(* IEC 61131-3 sources: 2026_Projet_YGO_ExcavatriceDragage/TOOLS/TEST_AUTO_CI/RESULTS/B_AU_SECURITE/tests/contract_deferred, 1 file *)

(* ---- test_fb_safety_emergency_contract_deferred.st ---- *)
(* Essais différés : causes, diagnostics et latches. Non exécutés par run.bat ; à reprendre dans le futur socle de contrat FB. *)
SETUP
VAR
    fb : FB_SAFETY_EMERGENCYMANAGEMENT;
END_VAR
END_SETUP

(* Ce fichier est volontairement hors execution run.bat. Migration prevue vers le socle de contrat FB. *)

TEST 'TC-P01-023 Etape invalide -> abandon trace et lockout'
    fb(ENABLE := TRUE, RESET := FALSE, ARMREQUEST := FALSE, POWERCUTOFFREQUEST := FALSE,
       BTNEMERGENCYCUTOFF := FALSE, EMERGENCYCHAINCLOSED := TRUE, POWERCONTACTORENGAGED := FALSE);
    fb(ENABLE := TRUE, RESET := FALSE, ARMREQUEST := FALSE, POWERCUTOFFREQUEST := FALSE,
       BTNEMERGENCYCUTOFF := FALSE, EMERGENCYCHAINCLOSED := TRUE, POWERCONTACTORENGAGED := FALSE);

    fb.ARMINGSEQSTEP := 7;
    ADVANCE_TIME(10000000);
    fb(ENABLE := TRUE, RESET := FALSE, ARMREQUEST := FALSE, POWERCUTOFFREQUEST := FALSE,
       BTNEMERGENCYCUTOFF := FALSE, EMERGENCYCHAINCLOSED := TRUE, POWERCONTACTORENGAGED := FALSE);
    fb(ENABLE := TRUE, RESET := FALSE, ARMREQUEST := FALSE, POWERCUTOFFREQUEST := FALSE,
       BTNEMERGENCYCUTOFF := FALSE, EMERGENCYCHAINCLOSED := TRUE, POWERCONTACTORENGAGED := FALSE);

    ASSERT_EQ(fb.STATUS.STATE.STEP, 0, 'etape inconnue -> IDLE');
    ASSERT_EQ(fb.STATUS.DIAG.LASTABORTSTEP, 7, 'etape inconnue tracee');
    ASSERT_EQ(fb.STATUS.DIAG.LASTABORTCAUSE, 256, 'cause = CST_ABORT_INVALID_STEP');
    ASSERT_TRUE(fb.STATUS.DIAG.LOCKOUTACTIVE, 'etape inconnue -> lockout');
    ASSERT_FALSE(fb.CMD.ARMPULSE_CMD, 'etape inconnue -> aucune impulsion');
    ASSERT_EQ(fb.STATUS.OPERATORMESSAGE, 'AU: etape sequence invalide - verifier puis Reset', 'etape inconnue -> message explicite');
END_TEST

TEST 'TC-P01-011 PowerCutOffRequest pendant l impulsion (step 5) -> abandon 16#0010 + lockout + Error=FALSE'
    (* Montee nominale jusqu au pulse (step 5), comme TC-P01-003 *)
    fb(ENABLE := TRUE, RESET := FALSE, ARMREQUEST := FALSE, POWERCUTOFFREQUEST := FALSE,
       BTNEMERGENCYCUTOFF := FALSE, EMERGENCYCHAINCLOSED := TRUE, POWERCONTACTORENGAGED := FALSE);
    fb(ENABLE := TRUE, RESET := FALSE, ARMREQUEST := FALSE, POWERCUTOFFREQUEST := FALSE,
       BTNEMERGENCYCUTOFF := FALSE, EMERGENCYCHAINCLOSED := TRUE, POWERCONTACTORENGAGED := FALSE);
    ADVANCE_TIME(10000000);
    fb(ENABLE := TRUE, RESET := FALSE, ARMREQUEST := FALSE, POWERCUTOFFREQUEST := FALSE,
       BTNEMERGENCYCUTOFF := FALSE, EMERGENCYCHAINCLOSED := TRUE, POWERCONTACTORENGAGED := FALSE);
    fb(ENABLE := TRUE, RESET := FALSE, ARMREQUEST := FALSE, POWERCUTOFFREQUEST := FALSE,
       BTNEMERGENCYCUTOFF := FALSE, EMERGENCYCHAINCLOSED := TRUE, POWERCONTACTORENGAGED := FALSE);
    ADVANCE_TIME(10000000);
    fb(ENABLE := TRUE, RESET := FALSE, ARMREQUEST := TRUE, POWERCUTOFFREQUEST := FALSE,
       BTNEMERGENCYCUTOFF := FALSE, EMERGENCYCHAINCLOSED := TRUE, POWERCONTACTORENGAGED := FALSE);
    fb(ENABLE := TRUE, RESET := FALSE, ARMREQUEST := TRUE, POWERCUTOFFREQUEST := FALSE,
       BTNEMERGENCYCUTOFF := FALSE, EMERGENCYCHAINCLOSED := TRUE, POWERCONTACTORENGAGED := FALSE);
    ADVANCE_TIME(200000000);
    fb(ENABLE := TRUE, RESET := FALSE, ARMREQUEST := FALSE, POWERCUTOFFREQUEST := FALSE,
       BTNEMERGENCYCUTOFF := FALSE, EMERGENCYCHAINCLOSED := FALSE, POWERCONTACTORENGAGED := FALSE);
    fb(ENABLE := TRUE, RESET := FALSE, ARMREQUEST := FALSE, POWERCUTOFFREQUEST := FALSE,
       BTNEMERGENCYCUTOFF := FALSE, EMERGENCYCHAINCLOSED := FALSE, POWERCONTACTORENGAGED := FALSE);
    ADVANCE_TIME(200000000);
    fb(ENABLE := TRUE, RESET := FALSE, ARMREQUEST := FALSE, POWERCUTOFFREQUEST := FALSE,
       BTNEMERGENCYCUTOFF := FALSE, EMERGENCYCHAINCLOSED := TRUE, POWERCONTACTORENGAGED := FALSE);
    fb(ENABLE := TRUE, RESET := FALSE, ARMREQUEST := FALSE, POWERCUTOFFREQUEST := FALSE,
       BTNEMERGENCYCUTOFF := FALSE, EMERGENCYCHAINCLOSED := TRUE, POWERCONTACTORENGAGED := FALSE);
    ADVANCE_TIME(200000000);
    fb(ENABLE := TRUE, RESET := FALSE, ARMREQUEST := FALSE, POWERCUTOFFREQUEST := FALSE,
       BTNEMERGENCYCUTOFF := FALSE, EMERGENCYCHAINCLOSED := FALSE, POWERCONTACTORENGAGED := FALSE);
    fb(ENABLE := TRUE, RESET := FALSE, ARMREQUEST := FALSE, POWERCUTOFFREQUEST := FALSE,
       BTNEMERGENCYCUTOFF := FALSE, EMERGENCYCHAINCLOSED := FALSE, POWERCONTACTORENGAGED := FALSE);
    ADVANCE_TIME(200000000);
    fb(ENABLE := TRUE, RESET := FALSE, ARMREQUEST := FALSE, POWERCUTOFFREQUEST := FALSE,
       BTNEMERGENCYCUTOFF := FALSE, EMERGENCYCHAINCLOSED := TRUE, POWERCONTACTORENGAGED := FALSE);
    fb(ENABLE := TRUE, RESET := FALSE, ARMREQUEST := FALSE, POWERCUTOFFREQUEST := FALSE,
       BTNEMERGENCYCUTOFF := FALSE, EMERGENCYCHAINCLOSED := TRUE, POWERCONTACTORENGAGED := FALSE);
    ASSERT_EQ(fb.STATUS.STATE.STEP, 5, 'les 2 canaux valides -> pulse (step 5)');
    ASSERT_TRUE(fb.CMD.ARMPULSE_CMD, 'precondition : pulse actif');

    (* Coupure metier PowerCutOffRequest PENDANT l impulsion (step 5) *)
    ADVANCE_TIME(10000000);
    fb(ENABLE := TRUE, RESET := FALSE, ARMREQUEST := FALSE, POWERCUTOFFREQUEST := TRUE,
       BTNEMERGENCYCUTOFF := FALSE, EMERGENCYCHAINCLOSED := TRUE, POWERCONTACTORENGAGED := FALSE);
    fb(ENABLE := TRUE, RESET := FALSE, ARMREQUEST := FALSE, POWERCUTOFFREQUEST := TRUE,
       BTNEMERGENCYCUTOFF := FALSE, EMERGENCYCHAINCLOSED := TRUE, POWERCONTACTORENGAGED := FALSE);
    ASSERT_EQ(fb.STATUS.STATE.STEP, 0, 'PowerCutOff pendant pulse -> sequence ramenee a IDLE');
    ASSERT_EQ(fb.STATUS.DIAG.LASTABORTCAUSE, 16#0010, 'cause abandon = 16#0010 (PowerCutOff metier)');
    ASSERT_EQ(fb.STATUS.DIAG.LASTABORTSTEP, 5, 'abandon a l etape 5 (impulsion)');
    ASSERT_TRUE(fb.STATUS.DIAG.LOCKOUTACTIVE, 'lockout 5s actif apres coupure metier');
    ASSERT_FALSE(fb.STATUS.DIAG.ERROR, 'coupure metier voulue -> PAS de defaut d armement (Error=FALSE)');
    ASSERT_FALSE(fb.STATUS.STATE.ARMABLE, 'interlock : PowerCutOffRequest actif -> Armable=FALSE');
    ASSERT_EQ(fb.STATUS.OPERATORMESSAGE, 'AU: coupure securite metier active - lever la cause puis rearmer', 'message coupure metier (priorite §11 sur le CASE)');
END_TEST

TEST 'TC-P01-012 Armable=1 mais rearmement echoue a l etape 5 (PowerCutOff pendant pulse)'
    (* Precondition : au repos boucle saine, Armable=TRUE (rearmement autorise) *)
    fb(ENABLE := TRUE, RESET := FALSE, ARMREQUEST := FALSE, POWERCUTOFFREQUEST := FALSE,
       BTNEMERGENCYCUTOFF := FALSE, EMERGENCYCHAINCLOSED := TRUE, POWERCONTACTORENGAGED := FALSE);
    fb(ENABLE := TRUE, RESET := FALSE, ARMREQUEST := FALSE, POWERCUTOFFREQUEST := FALSE,
       BTNEMERGENCYCUTOFF := FALSE, EMERGENCYCHAINCLOSED := TRUE, POWERCONTACTORENGAGED := FALSE);
    ADVANCE_TIME(10000000);
    fb(ENABLE := TRUE, RESET := FALSE, ARMREQUEST := FALSE, POWERCUTOFFREQUEST := FALSE,
       BTNEMERGENCYCUTOFF := FALSE, EMERGENCYCHAINCLOSED := TRUE, POWERCONTACTORENGAGED := FALSE);
    fb(ENABLE := TRUE, RESET := FALSE, ARMREQUEST := FALSE, POWERCUTOFFREQUEST := FALSE,
       BTNEMERGENCYCUTOFF := FALSE, EMERGENCYCHAINCLOSED := TRUE, POWERCONTACTORENGAGED := FALSE);
    ASSERT_TRUE(fb.STATUS.STATE.ARMABLE, 'precondition : Armable=TRUE (rearmement autorise)');

    (* Rearmement lance -> sequence demarre *)
    ADVANCE_TIME(10000000);
    fb(ENABLE := TRUE, RESET := FALSE, ARMREQUEST := TRUE, POWERCUTOFFREQUEST := FALSE,
       BTNEMERGENCYCUTOFF := FALSE, EMERGENCYCHAINCLOSED := TRUE, POWERCONTACTORENGAGED := FALSE);
    fb(ENABLE := TRUE, RESET := FALSE, ARMREQUEST := TRUE, POWERCUTOFFREQUEST := FALSE,
       BTNEMERGENCYCUTOFF := FALSE, EMERGENCYCHAINCLOSED := TRUE, POWERCONTACTORENGAGED := FALSE);
    ASSERT_EQ(fb.STATUS.STATE.STEP, 1, 'ArmRequest -> sequence lancee (step 1)');

    (* Montee nominale jusqu au pulse (step 5) *)
    ADVANCE_TIME(200000000);
    fb(ENABLE := TRUE, RESET := FALSE, ARMREQUEST := FALSE, POWERCUTOFFREQUEST := FALSE,
       BTNEMERGENCYCUTOFF := FALSE, EMERGENCYCHAINCLOSED := FALSE, POWERCONTACTORENGAGED := FALSE);
    fb(ENABLE := TRUE, RESET := FALSE, ARMREQUEST := FALSE, POWERCUTOFFREQUEST := FALSE,
       BTNEMERGENCYCUTOFF := FALSE, EMERGENCYCHAINCLOSED := FALSE, POWERCONTACTORENGAGED := FALSE);
    ADVANCE_TIME(200000000);
    fb(ENABLE := TRUE, RESET := FALSE, ARMREQUEST := FALSE, POWERCUTOFFREQUEST := FALSE,
       BTNEMERGENCYCUTOFF := FALSE, EMERGENCYCHAINCLOSED := TRUE, POWERCONTACTORENGAGED := FALSE);
    fb(ENABLE := TRUE, RESET := FALSE, ARMREQUEST := FALSE, POWERCUTOFFREQUEST := FALSE,
       BTNEMERGENCYCUTOFF := FALSE, EMERGENCYCHAINCLOSED := TRUE, POWERCONTACTORENGAGED := FALSE);
    ADVANCE_TIME(200000000);
    fb(ENABLE := TRUE, RESET := FALSE, ARMREQUEST := FALSE, POWERCUTOFFREQUEST := FALSE,
       BTNEMERGENCYCUTOFF := FALSE, EMERGENCYCHAINCLOSED := FALSE, POWERCONTACTORENGAGED := FALSE);
    fb(ENABLE := TRUE, RESET := FALSE, ARMREQUEST := FALSE, POWERCUTOFFREQUEST := FALSE,
       BTNEMERGENCYCUTOFF := FALSE, EMERGENCYCHAINCLOSED := FALSE, POWERCONTACTORENGAGED := FALSE);
    ADVANCE_TIME(200000000);
    fb(ENABLE := TRUE, RESET := FALSE, ARMREQUEST := FALSE, POWERCUTOFFREQUEST := FALSE,
       BTNEMERGENCYCUTOFF := FALSE, EMERGENCYCHAINCLOSED := TRUE, POWERCONTACTORENGAGED := FALSE);
    fb(ENABLE := TRUE, RESET := FALSE, ARMREQUEST := FALSE, POWERCUTOFFREQUEST := FALSE,
       BTNEMERGENCYCUTOFF := FALSE, EMERGENCYCHAINCLOSED := TRUE, POWERCONTACTORENGAGED := FALSE);
    ASSERT_EQ(fb.STATUS.STATE.STEP, 5, 'les 2 canaux valides -> pulse (step 5)');

    (* Coupure metier pendant l impulsion -> echec a l etape 5 *)
    ADVANCE_TIME(10000000);
    fb(ENABLE := TRUE, RESET := FALSE, ARMREQUEST := FALSE, POWERCUTOFFREQUEST := TRUE,
       BTNEMERGENCYCUTOFF := FALSE, EMERGENCYCHAINCLOSED := TRUE, POWERCONTACTORENGAGED := FALSE);
    fb(ENABLE := TRUE, RESET := FALSE, ARMREQUEST := FALSE, POWERCUTOFFREQUEST := TRUE,
       BTNEMERGENCYCUTOFF := FALSE, EMERGENCYCHAINCLOSED := TRUE, POWERCONTACTORENGAGED := FALSE);
    ASSERT_EQ(fb.STATUS.STATE.STEP, 0, 'echec a l etape 5 -> sequence ramenee a IDLE');
    ASSERT_EQ(fb.STATUS.DIAG.LASTABORTSTEP, 5, 'abandon a l etape 5');
    ASSERT_EQ(fb.STATUS.DIAG.LASTABORTCAUSE, 16#0010, 'cause = 16#0010 (PowerCutOff metier)');
    ASSERT_FALSE(fb.STATUS.DONE, 'rearmement NON abouti (Done=FALSE, contacteur non engage)');
    ASSERT_FALSE(fb.STATUS.DIAG.ERROR, 'echec silencieux : PAS de defaut d armement (Error=FALSE)');
END_TEST

TEST 'TC-P01-013 Recuperation Reset : cause latched -> Reset -> cause levee -> rearmement reussi'
    (* Montee nominale jusqu au pulse (step 5), puis coupure metier -> abandon 16#0010 + lockout *)
    fb(ENABLE := TRUE, RESET := FALSE, ARMREQUEST := FALSE, POWERCUTOFFREQUEST := FALSE,
       BTNEMERGENCYCUTOFF := FALSE, EMERGENCYCHAINCLOSED := TRUE, POWERCONTACTORENGAGED := FALSE);
    fb(ENABLE := TRUE, RESET := FALSE, ARMREQUEST := FALSE, POWERCUTOFFREQUEST := FALSE,
       BTNEMERGENCYCUTOFF := FALSE, EMERGENCYCHAINCLOSED := TRUE, POWERCONTACTORENGAGED := FALSE);
    ADVANCE_TIME(10000000);
    fb(ENABLE := TRUE, RESET := FALSE, ARMREQUEST := FALSE, POWERCUTOFFREQUEST := FALSE,
       BTNEMERGENCYCUTOFF := FALSE, EMERGENCYCHAINCLOSED := TRUE, POWERCONTACTORENGAGED := FALSE);
    fb(ENABLE := TRUE, RESET := FALSE, ARMREQUEST := FALSE, POWERCUTOFFREQUEST := FALSE,
       BTNEMERGENCYCUTOFF := FALSE, EMERGENCYCHAINCLOSED := TRUE, POWERCONTACTORENGAGED := FALSE);
    ADVANCE_TIME(10000000);
    fb(ENABLE := TRUE, RESET := FALSE, ARMREQUEST := TRUE, POWERCUTOFFREQUEST := FALSE,
       BTNEMERGENCYCUTOFF := FALSE, EMERGENCYCHAINCLOSED := TRUE, POWERCONTACTORENGAGED := FALSE);
    fb(ENABLE := TRUE, RESET := FALSE, ARMREQUEST := TRUE, POWERCUTOFFREQUEST := FALSE,
       BTNEMERGENCYCUTOFF := FALSE, EMERGENCYCHAINCLOSED := TRUE, POWERCONTACTORENGAGED := FALSE);
    ADVANCE_TIME(200000000);
    fb(ENABLE := TRUE, RESET := FALSE, ARMREQUEST := FALSE, POWERCUTOFFREQUEST := FALSE,
       BTNEMERGENCYCUTOFF := FALSE, EMERGENCYCHAINCLOSED := FALSE, POWERCONTACTORENGAGED := FALSE);
    fb(ENABLE := TRUE, RESET := FALSE, ARMREQUEST := FALSE, POWERCUTOFFREQUEST := FALSE,
       BTNEMERGENCYCUTOFF := FALSE, EMERGENCYCHAINCLOSED := FALSE, POWERCONTACTORENGAGED := FALSE);
    ADVANCE_TIME(200000000);
    fb(ENABLE := TRUE, RESET := FALSE, ARMREQUEST := FALSE, POWERCUTOFFREQUEST := FALSE,
       BTNEMERGENCYCUTOFF := FALSE, EMERGENCYCHAINCLOSED := TRUE, POWERCONTACTORENGAGED := FALSE);
    fb(ENABLE := TRUE, RESET := FALSE, ARMREQUEST := FALSE, POWERCUTOFFREQUEST := FALSE,
       BTNEMERGENCYCUTOFF := FALSE, EMERGENCYCHAINCLOSED := TRUE, POWERCONTACTORENGAGED := FALSE);
    ADVANCE_TIME(200000000);
    fb(ENABLE := TRUE, RESET := FALSE, ARMREQUEST := FALSE, POWERCUTOFFREQUEST := FALSE,
       BTNEMERGENCYCUTOFF := FALSE, EMERGENCYCHAINCLOSED := FALSE, POWERCONTACTORENGAGED := FALSE);
    fb(ENABLE := TRUE, RESET := FALSE, ARMREQUEST := FALSE, POWERCUTOFFREQUEST := FALSE,
       BTNEMERGENCYCUTOFF := FALSE, EMERGENCYCHAINCLOSED := FALSE, POWERCONTACTORENGAGED := FALSE);
    ADVANCE_TIME(200000000);
    fb(ENABLE := TRUE, RESET := FALSE, ARMREQUEST := FALSE, POWERCUTOFFREQUEST := FALSE,
       BTNEMERGENCYCUTOFF := FALSE, EMERGENCYCHAINCLOSED := TRUE, POWERCONTACTORENGAGED := FALSE);
    fb(ENABLE := TRUE, RESET := FALSE, ARMREQUEST := FALSE, POWERCUTOFFREQUEST := FALSE,
       BTNEMERGENCYCUTOFF := FALSE, EMERGENCYCHAINCLOSED := TRUE, POWERCONTACTORENGAGED := FALSE);
    ASSERT_EQ(fb.STATUS.STATE.STEP, 5, 'pulse (step 5)');

    (* Coupure metier -> abandon 16#0010 + lockout *)
    ADVANCE_TIME(10000000);
    fb(ENABLE := TRUE, RESET := FALSE, ARMREQUEST := FALSE, POWERCUTOFFREQUEST := TRUE,
       BTNEMERGENCYCUTOFF := FALSE, EMERGENCYCHAINCLOSED := TRUE, POWERCONTACTORENGAGED := FALSE);
    fb(ENABLE := TRUE, RESET := FALSE, ARMREQUEST := FALSE, POWERCUTOFFREQUEST := TRUE,
       BTNEMERGENCYCUTOFF := FALSE, EMERGENCYCHAINCLOSED := TRUE, POWERCONTACTORENGAGED := FALSE);
    ASSERT_EQ(fb.STATUS.DIAG.LASTABORTCAUSE, 16#0010, 'cause latched = 16#0010');
    ASSERT_TRUE(fb.STATUS.DIAG.LOCKOUTACTIVE, 'lockout actif');

    (* Cause levee (PowerCutOffRequest=FALSE) + Reset -> lockout purge, Armable redevient TRUE *)
    ADVANCE_TIME(10000000);
    fb(ENABLE := TRUE, RESET := TRUE, ARMREQUEST := FALSE, POWERCUTOFFREQUEST := FALSE,
       BTNEMERGENCYCUTOFF := FALSE, EMERGENCYCHAINCLOSED := TRUE, POWERCONTACTORENGAGED := FALSE);
    fb(ENABLE := TRUE, RESET := TRUE, ARMREQUEST := FALSE, POWERCUTOFFREQUEST := FALSE,
       BTNEMERGENCYCUTOFF := FALSE, EMERGENCYCHAINCLOSED := TRUE, POWERCONTACTORENGAGED := FALSE);
    ASSERT_FALSE(fb.STATUS.DIAG.LOCKOUTACTIVE, 'Reset purge le lockout');
    ASSERT_TRUE(fb.STATUS.STATE.ARMABLE, 'cause levee + Reset -> Armable=TRUE');

    (* Nouveau rearmement -> reussite (contacteur engage) *)
    ADVANCE_TIME(10000000);
    fb(ENABLE := TRUE, RESET := FALSE, ARMREQUEST := TRUE, POWERCUTOFFREQUEST := FALSE,
       BTNEMERGENCYCUTOFF := FALSE, EMERGENCYCHAINCLOSED := TRUE, POWERCONTACTORENGAGED := FALSE);
    fb(ENABLE := TRUE, RESET := FALSE, ARMREQUEST := TRUE, POWERCUTOFFREQUEST := FALSE,
       BTNEMERGENCYCUTOFF := FALSE, EMERGENCYCHAINCLOSED := TRUE, POWERCONTACTORENGAGED := FALSE);
    ASSERT_EQ(fb.STATUS.STATE.STEP, 1, 'nouveau front ArmRequest -> sequence relancee');
    ADVANCE_TIME(200000000);
    fb(ENABLE := TRUE, RESET := FALSE, ARMREQUEST := FALSE, POWERCUTOFFREQUEST := FALSE,
       BTNEMERGENCYCUTOFF := FALSE, EMERGENCYCHAINCLOSED := FALSE, POWERCONTACTORENGAGED := FALSE);
    fb(ENABLE := TRUE, RESET := FALSE, ARMREQUEST := FALSE, POWERCUTOFFREQUEST := FALSE,
       BTNEMERGENCYCUTOFF := FALSE, EMERGENCYCHAINCLOSED := FALSE, POWERCONTACTORENGAGED := FALSE);
    ADVANCE_TIME(200000000);
    fb(ENABLE := TRUE, RESET := FALSE, ARMREQUEST := FALSE, POWERCUTOFFREQUEST := FALSE,
       BTNEMERGENCYCUTOFF := FALSE, EMERGENCYCHAINCLOSED := TRUE, POWERCONTACTORENGAGED := FALSE);
    fb(ENABLE := TRUE, RESET := FALSE, ARMREQUEST := FALSE, POWERCUTOFFREQUEST := FALSE,
       BTNEMERGENCYCUTOFF := FALSE, EMERGENCYCHAINCLOSED := TRUE, POWERCONTACTORENGAGED := FALSE);
    ADVANCE_TIME(200000000);
    fb(ENABLE := TRUE, RESET := FALSE, ARMREQUEST := FALSE, POWERCUTOFFREQUEST := FALSE,
       BTNEMERGENCYCUTOFF := FALSE, EMERGENCYCHAINCLOSED := FALSE, POWERCONTACTORENGAGED := FALSE);
    fb(ENABLE := TRUE, RESET := FALSE, ARMREQUEST := FALSE, POWERCUTOFFREQUEST := FALSE,
       BTNEMERGENCYCUTOFF := FALSE, EMERGENCYCHAINCLOSED := FALSE, POWERCONTACTORENGAGED := FALSE);
    ADVANCE_TIME(200000000);
    fb(ENABLE := TRUE, RESET := FALSE, ARMREQUEST := FALSE, POWERCUTOFFREQUEST := FALSE,
       BTNEMERGENCYCUTOFF := FALSE, EMERGENCYCHAINCLOSED := TRUE, POWERCONTACTORENGAGED := FALSE);
    fb(ENABLE := TRUE, RESET := FALSE, ARMREQUEST := FALSE, POWERCUTOFFREQUEST := FALSE,
       BTNEMERGENCYCUTOFF := FALSE, EMERGENCYCHAINCLOSED := TRUE, POWERCONTACTORENGAGED := FALSE);
    ADVANCE_TIME(1000000000);
    fb(ENABLE := TRUE, RESET := FALSE, ARMREQUEST := FALSE, POWERCUTOFFREQUEST := FALSE,
       BTNEMERGENCYCUTOFF := FALSE, EMERGENCYCHAINCLOSED := TRUE, POWERCONTACTORENGAGED := FALSE);
    fb(ENABLE := TRUE, RESET := FALSE, ARMREQUEST := FALSE, POWERCUTOFFREQUEST := FALSE,
       BTNEMERGENCYCUTOFF := FALSE, EMERGENCYCHAINCLOSED := TRUE, POWERCONTACTORENGAGED := FALSE);
    ASSERT_EQ(fb.STATUS.STATE.STEP, 6, 'pulse termine -> attente confirmation');
    ADVANCE_TIME(10000000);
    fb(ENABLE := TRUE, RESET := FALSE, ARMREQUEST := FALSE, POWERCUTOFFREQUEST := FALSE,
       BTNEMERGENCYCUTOFF := FALSE, EMERGENCYCHAINCLOSED := TRUE, POWERCONTACTORENGAGED := TRUE);
    fb(ENABLE := TRUE, RESET := FALSE, ARMREQUEST := FALSE, POWERCUTOFFREQUEST := FALSE,
       BTNEMERGENCYCUTOFF := FALSE, EMERGENCYCHAINCLOSED := TRUE, POWERCONTACTORENGAGED := TRUE);
    ASSERT_EQ(fb.STATUS.STATE.STEP, 0, 'contacteur confirme -> retour IDLE');
    ASSERT_TRUE(fb.STATUS.DONE, 'rearmement reussi (Done=TRUE)');
    ASSERT_FALSE(fb.STATUS.DIAG.ERROR, 'aucun defaut apres reussite');
END_TEST

TEST 'TC-P01-014 Defaillance redondance B : canal B colle pendant TestB -> abandon 16#0040'
    (* 💤 Setup : demarrage + regime etabli, sain (boucle fermee, contacteur repos) *)
    fb(ENABLE := TRUE, RESET := FALSE, ARMREQUEST := FALSE, POWERCUTOFFREQUEST := FALSE,
       BTNEMERGENCYCUTOFF := FALSE, EMERGENCYCHAINCLOSED := TRUE, POWERCONTACTORENGAGED := FALSE);
    fb(ENABLE := TRUE, RESET := FALSE, ARMREQUEST := FALSE, POWERCUTOFFREQUEST := FALSE,
       BTNEMERGENCYCUTOFF := FALSE, EMERGENCYCHAINCLOSED := TRUE, POWERCONTACTORENGAGED := FALSE);
    ADVANCE_TIME(10000000);
    fb(ENABLE := TRUE, RESET := FALSE, ARMREQUEST := FALSE, POWERCUTOFFREQUEST := FALSE,
       BTNEMERGENCYCUTOFF := FALSE, EMERGENCYCHAINCLOSED := TRUE, POWERCONTACTORENGAGED := FALSE);
    fb(ENABLE := TRUE, RESET := FALSE, ARMREQUEST := FALSE, POWERCUTOFFREQUEST := FALSE,
       BTNEMERGENCYCUTOFF := FALSE, EMERGENCYCHAINCLOSED := TRUE, POWERCONTACTORENGAGED := FALSE);

    (* 🚀 t=0 : front ArmRequest -> TestA (step 1) *)
    ADVANCE_TIME(10000000);
    fb(ENABLE := TRUE, RESET := FALSE, ARMREQUEST := TRUE, POWERCUTOFFREQUEST := FALSE,
       BTNEMERGENCYCUTOFF := FALSE, EMERGENCYCHAINCLOSED := TRUE, POWERCONTACTORENGAGED := FALSE);
    fb(ENABLE := TRUE, RESET := FALSE, ARMREQUEST := TRUE, POWERCUTOFFREQUEST := FALSE,
       BTNEMERGENCYCUTOFF := FALSE, EMERGENCYCHAINCLOSED := TRUE, POWERCONTACTORENGAGED := FALSE);
    ASSERT_EQ(fb.STATUS.STATE.STEP, 1, 'front ArmRequest -> TestA (step 1)');

    (* 🔍 t=200ms : TestA reussi (boucle tombe) -> RestoreA (step 2) *)
    ADVANCE_TIME(200000000);
    fb(ENABLE := TRUE, RESET := FALSE, ARMREQUEST := FALSE, POWERCUTOFFREQUEST := FALSE,
       BTNEMERGENCYCUTOFF := FALSE, EMERGENCYCHAINCLOSED := FALSE, POWERCONTACTORENGAGED := FALSE);
    fb(ENABLE := TRUE, RESET := FALSE, ARMREQUEST := FALSE, POWERCUTOFFREQUEST := FALSE,
       BTNEMERGENCYCUTOFF := FALSE, EMERGENCYCHAINCLOSED := FALSE, POWERCONTACTORENGAGED := FALSE);
    ASSERT_EQ(fb.STATUS.STATE.STEP, 2, 'TestA reussi -> RestoreA (step 2)');

    (* 🔍 t=400ms : RestoreA reussi (boucle refermee) -> TestB (step 3) *)
    ADVANCE_TIME(200000000);
    fb(ENABLE := TRUE, RESET := FALSE, ARMREQUEST := FALSE, POWERCUTOFFREQUEST := FALSE,
       BTNEMERGENCYCUTOFF := FALSE, EMERGENCYCHAINCLOSED := TRUE, POWERCONTACTORENGAGED := FALSE);
    fb(ENABLE := TRUE, RESET := FALSE, ARMREQUEST := FALSE, POWERCUTOFFREQUEST := FALSE,
       BTNEMERGENCYCUTOFF := FALSE, EMERGENCYCHAINCLOSED := TRUE, POWERCONTACTORENGAGED := FALSE);
    ASSERT_EQ(fb.STATUS.STATE.STEP, 3, 'RestoreA reussi -> TestB (step 3)');

    (* ⚠️ t=600ms : TestB -> canal B colle : boucle RESTE fermee apres 200ms -> defaut redondance B *)
    ADVANCE_TIME(200000000);
    fb(ENABLE := TRUE, RESET := FALSE, ARMREQUEST := FALSE, POWERCUTOFFREQUEST := FALSE,
       BTNEMERGENCYCUTOFF := FALSE, EMERGENCYCHAINCLOSED := TRUE, POWERCONTACTORENGAGED := FALSE);
    fb(ENABLE := TRUE, RESET := FALSE, ARMREQUEST := FALSE, POWERCUTOFFREQUEST := FALSE,
       BTNEMERGENCYCUTOFF := FALSE, EMERGENCYCHAINCLOSED := TRUE, POWERCONTACTORENGAGED := FALSE);
    ASSERT_EQ(fb.STATUS.STATE.STEP, 0, 'canal B colle -> retour IDLE');
    ASSERT_EQ(fb.STATUS.DIAG.LASTABORTSTEP, 3, 'abandon a l etape 3 (TestB)');
    ASSERT_EQ(fb.STATUS.DIAG.LASTABORTCAUSE, 16#0040, 'cause = 16#0040 (Redundancy B)');
    ASSERT_TRUE(fb.STATUS.DIAG.REDUNDANCYTESTFAILED, 'defaut redondance leve');
    ASSERT_TRUE(fb.STATUS.DIAG.ERROR, 'defaut visible sur Error');
    ASSERT_FALSE(fb.CMD.MAINTAINA_CMD, 'canal colle bloque le maintien A (interlock Cause brute)');
    ASSERT_FALSE(fb.CMD.MAINTAINB_CMD, 'canal colle bloque le maintien B (interlock Cause brute)');
END_TEST

TEST 'TC-P01-015 Timeout restauration A : boucle ne revient pas apres TestA -> abandon 16#0004'
    (* 💤 Setup : demarrage + regime etabli, sain *)
    fb(ENABLE := TRUE, RESET := FALSE, ARMREQUEST := FALSE, POWERCUTOFFREQUEST := FALSE,
       BTNEMERGENCYCUTOFF := FALSE, EMERGENCYCHAINCLOSED := TRUE, POWERCONTACTORENGAGED := FALSE);
    fb(ENABLE := TRUE, RESET := FALSE, ARMREQUEST := FALSE, POWERCUTOFFREQUEST := FALSE,
       BTNEMERGENCYCUTOFF := FALSE, EMERGENCYCHAINCLOSED := TRUE, POWERCONTACTORENGAGED := FALSE);
    ADVANCE_TIME(10000000);
    fb(ENABLE := TRUE, RESET := FALSE, ARMREQUEST := FALSE, POWERCUTOFFREQUEST := FALSE,
       BTNEMERGENCYCUTOFF := FALSE, EMERGENCYCHAINCLOSED := TRUE, POWERCONTACTORENGAGED := FALSE);
    fb(ENABLE := TRUE, RESET := FALSE, ARMREQUEST := FALSE, POWERCUTOFFREQUEST := FALSE,
       BTNEMERGENCYCUTOFF := FALSE, EMERGENCYCHAINCLOSED := TRUE, POWERCONTACTORENGAGED := FALSE);

    (* 🚀 t=0 : front ArmRequest -> TestA (step 1) *)
    ADVANCE_TIME(10000000);
    fb(ENABLE := TRUE, RESET := FALSE, ARMREQUEST := TRUE, POWERCUTOFFREQUEST := FALSE,
       BTNEMERGENCYCUTOFF := FALSE, EMERGENCYCHAINCLOSED := TRUE, POWERCONTACTORENGAGED := FALSE);
    fb(ENABLE := TRUE, RESET := FALSE, ARMREQUEST := TRUE, POWERCUTOFFREQUEST := FALSE,
       BTNEMERGENCYCUTOFF := FALSE, EMERGENCYCHAINCLOSED := TRUE, POWERCONTACTORENGAGED := FALSE);
    ASSERT_EQ(fb.STATUS.STATE.STEP, 1, 'front ArmRequest -> TestA (step 1)');

    (* 🔍 t=200ms : TestA reussi (boucle tombe) -> RestoreA (step 2) *)
    ADVANCE_TIME(200000000);
    fb(ENABLE := TRUE, RESET := FALSE, ARMREQUEST := FALSE, POWERCUTOFFREQUEST := FALSE,
       BTNEMERGENCYCUTOFF := FALSE, EMERGENCYCHAINCLOSED := FALSE, POWERCONTACTORENGAGED := FALSE);
    fb(ENABLE := TRUE, RESET := FALSE, ARMREQUEST := FALSE, POWERCUTOFFREQUEST := FALSE,
       BTNEMERGENCYCUTOFF := FALSE, EMERGENCYCHAINCLOSED := FALSE, POWERCONTACTORENGAGED := FALSE);
    ASSERT_EQ(fb.STATUS.STATE.STEP, 2, 'TestA reussi -> RestoreA (step 2)');

    (* ⚠️ t=400ms : RestoreA timeout -> boucle ne revient PAS apres 200ms -> abandon 16#0004 *)
    ADVANCE_TIME(200000000);
    fb(ENABLE := TRUE, RESET := FALSE, ARMREQUEST := FALSE, POWERCUTOFFREQUEST := FALSE,
       BTNEMERGENCYCUTOFF := FALSE, EMERGENCYCHAINCLOSED := FALSE, POWERCONTACTORENGAGED := FALSE);
    fb(ENABLE := TRUE, RESET := FALSE, ARMREQUEST := FALSE, POWERCUTOFFREQUEST := FALSE,
       BTNEMERGENCYCUTOFF := FALSE, EMERGENCYCHAINCLOSED := FALSE, POWERCONTACTORENGAGED := FALSE);
    ASSERT_EQ(fb.STATUS.STATE.STEP, 0, 'timeout restauration A -> retour IDLE');
    ASSERT_EQ(fb.STATUS.DIAG.LASTABORTSTEP, 2, 'abandon a l etape 2 (RestoreA)');
    ASSERT_EQ(fb.STATUS.DIAG.LASTABORTCAUSE, 16#0004, 'cause = 16#0004 (Timeout Restore A)');
    ASSERT_FALSE(fb.STATUS.DIAG.ERROR, 'timeout restauration -> PAS de defaut d armement (Error=FALSE)');
    ASSERT_FALSE(fb.STATUS.DIAG.LOCKOUTACTIVE, 'timeout restauration -> PAS de lockout');
END_TEST

TEST 'TC-P01-016 Timeout restauration B : boucle ne revient pas apres TestB -> abandon 16#0008'
    (* 💤 Setup : demarrage + regime etabli, sain *)
    fb(ENABLE := TRUE, RESET := FALSE, ARMREQUEST := FALSE, POWERCUTOFFREQUEST := FALSE,
       BTNEMERGENCYCUTOFF := FALSE, EMERGENCYCHAINCLOSED := TRUE, POWERCONTACTORENGAGED := FALSE);
    fb(ENABLE := TRUE, RESET := FALSE, ARMREQUEST := FALSE, POWERCUTOFFREQUEST := FALSE,
       BTNEMERGENCYCUTOFF := FALSE, EMERGENCYCHAINCLOSED := TRUE, POWERCONTACTORENGAGED := FALSE);
    ADVANCE_TIME(10000000);
    fb(ENABLE := TRUE, RESET := FALSE, ARMREQUEST := FALSE, POWERCUTOFFREQUEST := FALSE,
       BTNEMERGENCYCUTOFF := FALSE, EMERGENCYCHAINCLOSED := TRUE, POWERCONTACTORENGAGED := FALSE);
    fb(ENABLE := TRUE, RESET := FALSE, ARMREQUEST := FALSE, POWERCUTOFFREQUEST := FALSE,
       BTNEMERGENCYCUTOFF := FALSE, EMERGENCYCHAINCLOSED := TRUE, POWERCONTACTORENGAGED := FALSE);

    (* 🚀 t=0 : front ArmRequest -> TestA (step 1) *)
    ADVANCE_TIME(10000000);
    fb(ENABLE := TRUE, RESET := FALSE, ARMREQUEST := TRUE, POWERCUTOFFREQUEST := FALSE,
       BTNEMERGENCYCUTOFF := FALSE, EMERGENCYCHAINCLOSED := TRUE, POWERCONTACTORENGAGED := FALSE);
    fb(ENABLE := TRUE, RESET := FALSE, ARMREQUEST := TRUE, POWERCUTOFFREQUEST := FALSE,
       BTNEMERGENCYCUTOFF := FALSE, EMERGENCYCHAINCLOSED := TRUE, POWERCONTACTORENGAGED := FALSE);
    (* 🔍 t=200ms : TestA -> RestoreA *)
    ADVANCE_TIME(200000000);
    fb(ENABLE := TRUE, RESET := FALSE, ARMREQUEST := FALSE, POWERCUTOFFREQUEST := FALSE,
       BTNEMERGENCYCUTOFF := FALSE, EMERGENCYCHAINCLOSED := FALSE, POWERCONTACTORENGAGED := FALSE);
    fb(ENABLE := TRUE, RESET := FALSE, ARMREQUEST := FALSE, POWERCUTOFFREQUEST := FALSE,
       BTNEMERGENCYCUTOFF := FALSE, EMERGENCYCHAINCLOSED := FALSE, POWERCONTACTORENGAGED := FALSE);
    (* 🔍 t=400ms : RestoreA -> TestB *)
    ADVANCE_TIME(200000000);
    fb(ENABLE := TRUE, RESET := FALSE, ARMREQUEST := FALSE, POWERCUTOFFREQUEST := FALSE,
       BTNEMERGENCYCUTOFF := FALSE, EMERGENCYCHAINCLOSED := TRUE, POWERCONTACTORENGAGED := FALSE);
    fb(ENABLE := TRUE, RESET := FALSE, ARMREQUEST := FALSE, POWERCUTOFFREQUEST := FALSE,
       BTNEMERGENCYCUTOFF := FALSE, EMERGENCYCHAINCLOSED := TRUE, POWERCONTACTORENGAGED := FALSE);
    (* 🔍 t=600ms : TestB -> RestoreB *)
    ADVANCE_TIME(200000000);
    fb(ENABLE := TRUE, RESET := FALSE, ARMREQUEST := FALSE, POWERCUTOFFREQUEST := FALSE,
       BTNEMERGENCYCUTOFF := FALSE, EMERGENCYCHAINCLOSED := FALSE, POWERCONTACTORENGAGED := FALSE);
    fb(ENABLE := TRUE, RESET := FALSE, ARMREQUEST := FALSE, POWERCUTOFFREQUEST := FALSE,
       BTNEMERGENCYCUTOFF := FALSE, EMERGENCYCHAINCLOSED := FALSE, POWERCONTACTORENGAGED := FALSE);
    ASSERT_EQ(fb.STATUS.STATE.STEP, 4, 'TestB reussi -> RestoreB (step 4)');

    (* ⚠️ t=800ms : RestoreB timeout -> boucle ne revient PAS apres 200ms -> abandon 16#0008 *)
    ADVANCE_TIME(200000000);
    fb(ENABLE := TRUE, RESET := FALSE, ARMREQUEST := FALSE, POWERCUTOFFREQUEST := FALSE,
       BTNEMERGENCYCUTOFF := FALSE, EMERGENCYCHAINCLOSED := FALSE, POWERCONTACTORENGAGED := FALSE);
    fb(ENABLE := TRUE, RESET := FALSE, ARMREQUEST := FALSE, POWERCUTOFFREQUEST := FALSE,
       BTNEMERGENCYCUTOFF := FALSE, EMERGENCYCHAINCLOSED := FALSE, POWERCONTACTORENGAGED := FALSE);
    ASSERT_EQ(fb.STATUS.STATE.STEP, 0, 'timeout restauration B -> retour IDLE');
    ASSERT_EQ(fb.STATUS.DIAG.LASTABORTSTEP, 4, 'abandon a l etape 4 (RestoreB)');
    ASSERT_EQ(fb.STATUS.DIAG.LASTABORTCAUSE, 16#0008, 'cause = 16#0008 (Timeout Restore B)');
    ASSERT_FALSE(fb.STATUS.DIAG.ERROR, 'timeout restauration B -> PAS de defaut d armement (Error=FALSE)');
    ASSERT_FALSE(fb.STATUS.DIAG.LOCKOUTACTIVE, 'timeout restauration B -> PAS de lockout');
END_TEST

TEST 'TC-P01-017 Chute de boucle pendant PULSE (step 5) -> abandon 16#0002 + lockout'
    (* 💤 Setup : demarrage + regime etabli, sain *)
    fb(ENABLE := TRUE, RESET := FALSE, ARMREQUEST := FALSE, POWERCUTOFFREQUEST := FALSE,
       BTNEMERGENCYCUTOFF := FALSE, EMERGENCYCHAINCLOSED := TRUE, POWERCONTACTORENGAGED := FALSE);
    fb(ENABLE := TRUE, RESET := FALSE, ARMREQUEST := FALSE, POWERCUTOFFREQUEST := FALSE,
       BTNEMERGENCYCUTOFF := FALSE, EMERGENCYCHAINCLOSED := TRUE, POWERCONTACTORENGAGED := FALSE);
    ADVANCE_TIME(10000000);
    fb(ENABLE := TRUE, RESET := FALSE, ARMREQUEST := FALSE, POWERCUTOFFREQUEST := FALSE,
       BTNEMERGENCYCUTOFF := FALSE, EMERGENCYCHAINCLOSED := TRUE, POWERCONTACTORENGAGED := FALSE);
    fb(ENABLE := TRUE, RESET := FALSE, ARMREQUEST := FALSE, POWERCUTOFFREQUEST := FALSE,
       BTNEMERGENCYCUTOFF := FALSE, EMERGENCYCHAINCLOSED := TRUE, POWERCONTACTORENGAGED := FALSE);
    (* 🚀 t=0 : front ArmRequest -> TestA *)
    ADVANCE_TIME(10000000);
    fb(ENABLE := TRUE, RESET := FALSE, ARMREQUEST := TRUE, POWERCUTOFFREQUEST := FALSE,
       BTNEMERGENCYCUTOFF := FALSE, EMERGENCYCHAINCLOSED := TRUE, POWERCONTACTORENGAGED := FALSE);
    fb(ENABLE := TRUE, RESET := FALSE, ARMREQUEST := TRUE, POWERCUTOFFREQUEST := FALSE,
       BTNEMERGENCYCUTOFF := FALSE, EMERGENCYCHAINCLOSED := TRUE, POWERCONTACTORENGAGED := FALSE);
    (* 🔍 t=200ms : TestA -> RestoreA *)
    ADVANCE_TIME(200000000);
    fb(ENABLE := TRUE, RESET := FALSE, ARMREQUEST := FALSE, POWERCUTOFFREQUEST := FALSE,
       BTNEMERGENCYCUTOFF := FALSE, EMERGENCYCHAINCLOSED := FALSE, POWERCONTACTORENGAGED := FALSE);
    fb(ENABLE := TRUE, RESET := FALSE, ARMREQUEST := FALSE, POWERCUTOFFREQUEST := FALSE,
       BTNEMERGENCYCUTOFF := FALSE, EMERGENCYCHAINCLOSED := FALSE, POWERCONTACTORENGAGED := FALSE);
    (* 🔍 t=400ms : RestoreA -> TestB *)
    ADVANCE_TIME(200000000);
    fb(ENABLE := TRUE, RESET := FALSE, ARMREQUEST := FALSE, POWERCUTOFFREQUEST := FALSE,
       BTNEMERGENCYCUTOFF := FALSE, EMERGENCYCHAINCLOSED := TRUE, POWERCONTACTORENGAGED := FALSE);
    fb(ENABLE := TRUE, RESET := FALSE, ARMREQUEST := FALSE, POWERCUTOFFREQUEST := FALSE,
       BTNEMERGENCYCUTOFF := FALSE, EMERGENCYCHAINCLOSED := TRUE, POWERCONTACTORENGAGED := FALSE);
    (* 🔍 t=600ms : TestB -> RestoreB *)
    ADVANCE_TIME(200000000);
    fb(ENABLE := TRUE, RESET := FALSE, ARMREQUEST := FALSE, POWERCUTOFFREQUEST := FALSE,
       BTNEMERGENCYCUTOFF := FALSE, EMERGENCYCHAINCLOSED := FALSE, POWERCONTACTORENGAGED := FALSE);
    fb(ENABLE := TRUE, RESET := FALSE, ARMREQUEST := FALSE, POWERCUTOFFREQUEST := FALSE,
       BTNEMERGENCYCUTOFF := FALSE, EMERGENCYCHAINCLOSED := FALSE, POWERCONTACTORENGAGED := FALSE);
    (* 🔍 t=800ms : RestoreB -> PULSE (step 5) *)
    ADVANCE_TIME(200000000);
    fb(ENABLE := TRUE, RESET := FALSE, ARMREQUEST := FALSE, POWERCUTOFFREQUEST := FALSE,
       BTNEMERGENCYCUTOFF := FALSE, EMERGENCYCHAINCLOSED := TRUE, POWERCONTACTORENGAGED := FALSE);
    fb(ENABLE := TRUE, RESET := FALSE, ARMREQUEST := FALSE, POWERCUTOFFREQUEST := FALSE,
       BTNEMERGENCYCUTOFF := FALSE, EMERGENCYCHAINCLOSED := TRUE, POWERCONTACTORENGAGED := FALSE);
    ASSERT_EQ(fb.STATUS.STATE.STEP, 5, 'les 2 canaux valides -> pulse (step 5)');
    ASSERT_TRUE(fb.CMD.ARMPULSE_CMD, 'precondition : pulse actif');

    (* ⚠️ t=810ms : chute de boucle materielle PENDANT l impulsion (step 5) *)
    ADVANCE_TIME(10000000);
    fb(ENABLE := TRUE, RESET := FALSE, ARMREQUEST := FALSE, POWERCUTOFFREQUEST := FALSE,
       BTNEMERGENCYCUTOFF := FALSE, EMERGENCYCHAINCLOSED := FALSE, POWERCONTACTORENGAGED := FALSE);
    fb(ENABLE := TRUE, RESET := FALSE, ARMREQUEST := FALSE, POWERCUTOFFREQUEST := FALSE,
       BTNEMERGENCYCUTOFF := FALSE, EMERGENCYCHAINCLOSED := FALSE, POWERCONTACTORENGAGED := FALSE);
    ASSERT_EQ(fb.STATUS.STATE.STEP, 0, 'chute boucle pendant pulse -> sequence ramenee a IDLE');
    ASSERT_EQ(fb.STATUS.DIAG.LASTABORTSTEP, 5, 'abandon a l etape 5 (pulse)');
    ASSERT_EQ(fb.STATUS.DIAG.LASTABORTCAUSE, 16#0002, 'cause = 16#0002 (Chute chaine)');
    ASSERT_TRUE(fb.STATUS.DIAG.ARMFAILED, 'chute boucle -> defaut EmergencyArmingFailed leve');
    ASSERT_TRUE(fb.STATUS.DIAG.LOCKOUTACTIVE, 'chute boucle -> lockout 5s actif');
    ASSERT_TRUE(fb.STATUS.DIAG.ERROR, 'defaut visible sur Error');
    ASSERT_FALSE(fb.CMD.ARMPULSE_CMD, 'pulse coupe immediatement');
END_TEST

TEST 'TC-P01-018 Chute de boucle pendant CONFIRM (step 6) -> abandon 16#0002 + lockout'
    (* 💤 Setup : demarrage + regime etabli, sain *)
    fb(ENABLE := TRUE, RESET := FALSE, ARMREQUEST := FALSE, POWERCUTOFFREQUEST := FALSE,
       BTNEMERGENCYCUTOFF := FALSE, EMERGENCYCHAINCLOSED := TRUE, POWERCONTACTORENGAGED := FALSE);
    fb(ENABLE := TRUE, RESET := FALSE, ARMREQUEST := FALSE, POWERCUTOFFREQUEST := FALSE,
       BTNEMERGENCYCUTOFF := FALSE, EMERGENCYCHAINCLOSED := TRUE, POWERCONTACTORENGAGED := FALSE);
    ADVANCE_TIME(10000000);
    fb(ENABLE := TRUE, RESET := FALSE, ARMREQUEST := FALSE, POWERCUTOFFREQUEST := FALSE,
       BTNEMERGENCYCUTOFF := FALSE, EMERGENCYCHAINCLOSED := TRUE, POWERCONTACTORENGAGED := FALSE);
    fb(ENABLE := TRUE, RESET := FALSE, ARMREQUEST := FALSE, POWERCUTOFFREQUEST := FALSE,
       BTNEMERGENCYCUTOFF := FALSE, EMERGENCYCHAINCLOSED := TRUE, POWERCONTACTORENGAGED := FALSE);
    (* 🚀 t=0 : front ArmRequest -> TestA *)
    ADVANCE_TIME(10000000);
    fb(ENABLE := TRUE, RESET := FALSE, ARMREQUEST := TRUE, POWERCUTOFFREQUEST := FALSE,
       BTNEMERGENCYCUTOFF := FALSE, EMERGENCYCHAINCLOSED := TRUE, POWERCONTACTORENGAGED := FALSE);
    fb(ENABLE := TRUE, RESET := FALSE, ARMREQUEST := TRUE, POWERCUTOFFREQUEST := FALSE,
       BTNEMERGENCYCUTOFF := FALSE, EMERGENCYCHAINCLOSED := TRUE, POWERCONTACTORENGAGED := FALSE);
    (* 🔍 t=200ms : TestA -> RestoreA *)
    ADVANCE_TIME(200000000);
    fb(ENABLE := TRUE, RESET := FALSE, ARMREQUEST := FALSE, POWERCUTOFFREQUEST := FALSE,
       BTNEMERGENCYCUTOFF := FALSE, EMERGENCYCHAINCLOSED := FALSE, POWERCONTACTORENGAGED := FALSE);
    fb(ENABLE := TRUE, RESET := FALSE, ARMREQUEST := FALSE, POWERCUTOFFREQUEST := FALSE,
       BTNEMERGENCYCUTOFF := FALSE, EMERGENCYCHAINCLOSED := FALSE, POWERCONTACTORENGAGED := FALSE);
    (* 🔍 t=400ms : RestoreA -> TestB *)
    ADVANCE_TIME(200000000);
    fb(ENABLE := TRUE, RESET := FALSE, ARMREQUEST := FALSE, POWERCUTOFFREQUEST := FALSE,
       BTNEMERGENCYCUTOFF := FALSE, EMERGENCYCHAINCLOSED := TRUE, POWERCONTACTORENGAGED := FALSE);
    fb(ENABLE := TRUE, RESET := FALSE, ARMREQUEST := FALSE, POWERCUTOFFREQUEST := FALSE,
       BTNEMERGENCYCUTOFF := FALSE, EMERGENCYCHAINCLOSED := TRUE, POWERCONTACTORENGAGED := FALSE);
    (* 🔍 t=600ms : TestB -> RestoreB *)
    ADVANCE_TIME(200000000);
    fb(ENABLE := TRUE, RESET := FALSE, ARMREQUEST := FALSE, POWERCUTOFFREQUEST := FALSE,
       BTNEMERGENCYCUTOFF := FALSE, EMERGENCYCHAINCLOSED := FALSE, POWERCONTACTORENGAGED := FALSE);
    fb(ENABLE := TRUE, RESET := FALSE, ARMREQUEST := FALSE, POWERCUTOFFREQUEST := FALSE,
       BTNEMERGENCYCUTOFF := FALSE, EMERGENCYCHAINCLOSED := FALSE, POWERCONTACTORENGAGED := FALSE);
    (* 🔍 t=800ms : RestoreB -> PULSE (step 5) *)
    ADVANCE_TIME(200000000);
    fb(ENABLE := TRUE, RESET := FALSE, ARMREQUEST := FALSE, POWERCUTOFFREQUEST := FALSE,
       BTNEMERGENCYCUTOFF := FALSE, EMERGENCYCHAINCLOSED := TRUE, POWERCONTACTORENGAGED := FALSE);
    fb(ENABLE := TRUE, RESET := FALSE, ARMREQUEST := FALSE, POWERCUTOFFREQUEST := FALSE,
       BTNEMERGENCYCUTOFF := FALSE, EMERGENCYCHAINCLOSED := TRUE, POWERCONTACTORENGAGED := FALSE);
    (* ⏱️ t=1.8s : pulse 1s termine -> CONFIRM (step 6) *)
    ADVANCE_TIME(1000000000);
    fb(ENABLE := TRUE, RESET := FALSE, ARMREQUEST := FALSE, POWERCUTOFFREQUEST := FALSE,
       BTNEMERGENCYCUTOFF := FALSE, EMERGENCYCHAINCLOSED := TRUE, POWERCONTACTORENGAGED := FALSE);
    fb(ENABLE := TRUE, RESET := FALSE, ARMREQUEST := FALSE, POWERCUTOFFREQUEST := FALSE,
       BTNEMERGENCYCUTOFF := FALSE, EMERGENCYCHAINCLOSED := TRUE, POWERCONTACTORENGAGED := FALSE);
    ASSERT_EQ(fb.STATUS.STATE.STEP, 6, 'pulse termine -> attente confirmation (step 6)');

    (* ⚠️ t=1.81s : chute de boucle materielle PENDANT la confirmation (step 6) *)
    ADVANCE_TIME(10000000);
    fb(ENABLE := TRUE, RESET := FALSE, ARMREQUEST := FALSE, POWERCUTOFFREQUEST := FALSE,
       BTNEMERGENCYCUTOFF := FALSE, EMERGENCYCHAINCLOSED := FALSE, POWERCONTACTORENGAGED := FALSE);
    fb(ENABLE := TRUE, RESET := FALSE, ARMREQUEST := FALSE, POWERCUTOFFREQUEST := FALSE,
       BTNEMERGENCYCUTOFF := FALSE, EMERGENCYCHAINCLOSED := FALSE, POWERCONTACTORENGAGED := FALSE);
    ASSERT_EQ(fb.STATUS.STATE.STEP, 0, 'chute boucle pendant confirm -> sequence ramenee a IDLE');
    ASSERT_EQ(fb.STATUS.DIAG.LASTABORTSTEP, 6, 'abandon a l etape 6 (confirm)');
    ASSERT_EQ(fb.STATUS.DIAG.LASTABORTCAUSE, 16#0002, 'cause = 16#0002 (Chute chaine)');
    ASSERT_TRUE(fb.STATUS.DIAG.ARMFAILED, 'chute boucle -> defaut EmergencyArmingFailed leve');
    ASSERT_TRUE(fb.STATUS.DIAG.LOCKOUTACTIVE, 'chute boucle -> lockout 5s actif');
    ASSERT_TRUE(fb.STATUS.DIAG.ERROR, 'defaut visible sur Error');
END_TEST

TEST 'TC-P01-019 Coupure IHM pendant la sequence -> abandon 16#0001 sans alarme ni lockout'
    (* 💤 Setup : demarrage + regime etabli, sain *)
    fb(ENABLE := TRUE, RESET := FALSE, ARMREQUEST := FALSE, POWERCUTOFFREQUEST := FALSE,
       BTNEMERGENCYCUTOFF := FALSE, EMERGENCYCHAINCLOSED := TRUE, POWERCONTACTORENGAGED := FALSE);
    fb(ENABLE := TRUE, RESET := FALSE, ARMREQUEST := FALSE, POWERCUTOFFREQUEST := FALSE,
       BTNEMERGENCYCUTOFF := FALSE, EMERGENCYCHAINCLOSED := TRUE, POWERCONTACTORENGAGED := FALSE);
    ADVANCE_TIME(10000000);
    fb(ENABLE := TRUE, RESET := FALSE, ARMREQUEST := FALSE, POWERCUTOFFREQUEST := FALSE,
       BTNEMERGENCYCUTOFF := FALSE, EMERGENCYCHAINCLOSED := TRUE, POWERCONTACTORENGAGED := FALSE);
    fb(ENABLE := TRUE, RESET := FALSE, ARMREQUEST := FALSE, POWERCUTOFFREQUEST := FALSE,
       BTNEMERGENCYCUTOFF := FALSE, EMERGENCYCHAINCLOSED := TRUE, POWERCONTACTORENGAGED := FALSE);
    (* 🚀 t=0 : front ArmRequest -> TestA *)
    ADVANCE_TIME(10000000);
    fb(ENABLE := TRUE, RESET := FALSE, ARMREQUEST := TRUE, POWERCUTOFFREQUEST := FALSE,
       BTNEMERGENCYCUTOFF := FALSE, EMERGENCYCHAINCLOSED := TRUE, POWERCONTACTORENGAGED := FALSE);
    fb(ENABLE := TRUE, RESET := FALSE, ARMREQUEST := TRUE, POWERCUTOFFREQUEST := FALSE,
       BTNEMERGENCYCUTOFF := FALSE, EMERGENCYCHAINCLOSED := TRUE, POWERCONTACTORENGAGED := FALSE);
    (* 🔍 t=200ms : TestA -> RestoreA *)
    ADVANCE_TIME(200000000);
    fb(ENABLE := TRUE, RESET := FALSE, ARMREQUEST := FALSE, POWERCUTOFFREQUEST := FALSE,
       BTNEMERGENCYCUTOFF := FALSE, EMERGENCYCHAINCLOSED := FALSE, POWERCONTACTORENGAGED := FALSE);
    fb(ENABLE := TRUE, RESET := FALSE, ARMREQUEST := FALSE, POWERCUTOFFREQUEST := FALSE,
       BTNEMERGENCYCUTOFF := FALSE, EMERGENCYCHAINCLOSED := FALSE, POWERCONTACTORENGAGED := FALSE);
    (* 🔍 t=400ms : RestoreA -> TestB *)
    ADVANCE_TIME(200000000);
    fb(ENABLE := TRUE, RESET := FALSE, ARMREQUEST := FALSE, POWERCUTOFFREQUEST := FALSE,
       BTNEMERGENCYCUTOFF := FALSE, EMERGENCYCHAINCLOSED := TRUE, POWERCONTACTORENGAGED := FALSE);
    fb(ENABLE := TRUE, RESET := FALSE, ARMREQUEST := FALSE, POWERCUTOFFREQUEST := FALSE,
       BTNEMERGENCYCUTOFF := FALSE, EMERGENCYCHAINCLOSED := TRUE, POWERCONTACTORENGAGED := FALSE);
    (* 🔍 t=600ms : TestB -> RestoreB *)
    ADVANCE_TIME(200000000);
    fb(ENABLE := TRUE, RESET := FALSE, ARMREQUEST := FALSE, POWERCUTOFFREQUEST := FALSE,
       BTNEMERGENCYCUTOFF := FALSE, EMERGENCYCHAINCLOSED := FALSE, POWERCONTACTORENGAGED := FALSE);
    fb(ENABLE := TRUE, RESET := FALSE, ARMREQUEST := FALSE, POWERCUTOFFREQUEST := FALSE,
       BTNEMERGENCYCUTOFF := FALSE, EMERGENCYCHAINCLOSED := FALSE, POWERCONTACTORENGAGED := FALSE);
    (* 🔍 t=800ms : RestoreB -> PULSE (step 5) *)
    ADVANCE_TIME(200000000);
    fb(ENABLE := TRUE, RESET := FALSE, ARMREQUEST := FALSE, POWERCUTOFFREQUEST := FALSE,
       BTNEMERGENCYCUTOFF := FALSE, EMERGENCYCHAINCLOSED := TRUE, POWERCONTACTORENGAGED := FALSE);
    fb(ENABLE := TRUE, RESET := FALSE, ARMREQUEST := FALSE, POWERCUTOFFREQUEST := FALSE,
       BTNEMERGENCYCUTOFF := FALSE, EMERGENCYCHAINCLOSED := TRUE, POWERCONTACTORENGAGED := FALSE);
    ASSERT_EQ(fb.STATUS.STATE.STEP, 5, 'les 2 canaux valides -> pulse (step 5)');

    (* 🛑 t=810ms : operateur appuie sur la coupure d urgence IHM PENDANT la sequence (step 5) *)
    ADVANCE_TIME(10000000);
    fb(ENABLE := TRUE, RESET := FALSE, ARMREQUEST := FALSE, POWERCUTOFFREQUEST := FALSE,
       BTNEMERGENCYCUTOFF := TRUE, EMERGENCYCHAINCLOSED := TRUE, POWERCONTACTORENGAGED := FALSE);
    fb(ENABLE := TRUE, RESET := FALSE, ARMREQUEST := FALSE, POWERCUTOFFREQUEST := FALSE,
       BTNEMERGENCYCUTOFF := TRUE, EMERGENCYCHAINCLOSED := TRUE, POWERCONTACTORENGAGED := FALSE);
    ASSERT_EQ(fb.STATUS.STATE.STEP, 0, 'coupure IHM -> sequence ramenee a IDLE');
    ASSERT_EQ(fb.STATUS.OPERATORMESSAGE, 'AU: coupure urgence IHM active - relacher puis rearmer', 'message coupure IHM (priorite §11 sur le CASE)');
    ASSERT_EQ(fb.STATUS.DIAG.LASTABORTSTEP, 5, 'abandon a l etape 5 (pulse)');
    ASSERT_EQ(fb.STATUS.DIAG.LASTABORTCAUSE, 16#0001, 'cause = 16#0001 (Cut IHM)');
    ASSERT_FALSE(fb.STATUS.DIAG.ERROR, 'coupure IHM volontaire -> PAS de defaut (Error=FALSE)');
    ASSERT_FALSE(fb.STATUS.DIAG.LOCKOUTACTIVE, 'coupure IHM volontaire -> PAS de lockout');
    ASSERT_FALSE(fb.CMD.ARMPULSE_CMD, 'pulse coupe immediatement');
    ASSERT_FALSE(fb.CMD.MAINTAINA_CMD, 'maintien A coupe');
    ASSERT_FALSE(fb.CMD.MAINTAINB_CMD, 'maintien B coupe');
END_TEST

TEST 'TC-P01-020 Autotest demarrage : chaine ouverte au 1er Enable -> StartupFail, Reset recupere'
    (* 🏁 t=0 : Enable=TRUE avec chaine AU OUVERTE -> autotest demarrage echoue (StartupFail) *)
    fb(ENABLE := TRUE, RESET := FALSE, ARMREQUEST := FALSE, POWERCUTOFFREQUEST := FALSE,
       BTNEMERGENCYCUTOFF := FALSE, EMERGENCYCHAINCLOSED := FALSE, POWERCONTACTORENGAGED := FALSE);
    fb(ENABLE := TRUE, RESET := FALSE, ARMREQUEST := FALSE, POWERCUTOFFREQUEST := FALSE,
       BTNEMERGENCYCUTOFF := FALSE, EMERGENCYCHAINCLOSED := FALSE, POWERCONTACTORENGAGED := FALSE);
    ASSERT_FALSE(fb.STATUS.READY, 'chaine ouverte au 1er Enable -> Ready=FALSE (StartupFail)');
    ASSERT_TRUE(fb.STATUS.DIAG.ERROR, 'autotest demarrage echoue -> Error=TRUE');
    ASSERT_EQ(fb.STATUS.OPERATORMESSAGE, 'AU: autotest demarrage echoue - verifier boucle/contacteur puis Reset', 'message autotest demarrage echoue (priorite §11)');
    ASSERT_EQ(fb.STATUS.DIAG.ERRORID, 16#0008, 'ErrorId bit3 = StartupFail (16#0008)');
    ASSERT_FALSE(fb.STATUS.STATE.ARMABLE, 'StartupFail -> Armable=FALSE');

    (* 🔄 t=10ms : chaine refermee mais StartupFail latche -> toujours pas Ready *)
    ADVANCE_TIME(10000000);
    fb(ENABLE := TRUE, RESET := FALSE, ARMREQUEST := FALSE, POWERCUTOFFREQUEST := FALSE,
       BTNEMERGENCYCUTOFF := FALSE, EMERGENCYCHAINCLOSED := TRUE, POWERCONTACTORENGAGED := FALSE);
    fb(ENABLE := TRUE, RESET := FALSE, ARMREQUEST := FALSE, POWERCUTOFFREQUEST := FALSE,
       BTNEMERGENCYCUTOFF := FALSE, EMERGENCYCHAINCLOSED := TRUE, POWERCONTACTORENGAGED := FALSE);
    ASSERT_FALSE(fb.STATUS.READY, 'StartupFail latche -> Ready reste FALSE meme chaine refermee');

    (* ✅ t=20ms : Reset -> StartupFail purge, Ready=TRUE *)
    ADVANCE_TIME(10000000);
    fb(ENABLE := TRUE, RESET := TRUE, ARMREQUEST := FALSE, POWERCUTOFFREQUEST := FALSE,
       BTNEMERGENCYCUTOFF := FALSE, EMERGENCYCHAINCLOSED := TRUE, POWERCONTACTORENGAGED := FALSE);
    fb(ENABLE := TRUE, RESET := TRUE, ARMREQUEST := FALSE, POWERCUTOFFREQUEST := FALSE,
       BTNEMERGENCYCUTOFF := FALSE, EMERGENCYCHAINCLOSED := TRUE, POWERCONTACTORENGAGED := FALSE);
    ASSERT_TRUE(fb.STATUS.READY, 'Reset purge StartupFail -> Ready=TRUE');
    ASSERT_FALSE(fb.STATUS.DIAG.ERROR, 'Reset acquitte le defaut -> Error=FALSE');
    ASSERT_TRUE(fb.STATUS.STATE.ARMABLE, 'apres Reset -> Armable=TRUE');
    ASSERT_EQ(fb.STATUS.OPERATORMESSAGE, 'AU: repos - pret a rearmer', 'message CASE 0/IDLE apres purge StartupFail par Reset');
END_TEST

TEST 'TC-P01-021 Enable=FALSE pendant l impulsion (step 5) -> neutralisation fail-safe immediate'
    (* 💤 t=-20ms : demarrage + regime etabli, sain (boucle fermee, contacteur repos) *)
    fb(ENABLE := TRUE, RESET := FALSE, ARMREQUEST := FALSE, POWERCUTOFFREQUEST := FALSE,
       BTNEMERGENCYCUTOFF := FALSE, EMERGENCYCHAINCLOSED := TRUE, POWERCONTACTORENGAGED := FALSE);
    fb(ENABLE := TRUE, RESET := FALSE, ARMREQUEST := FALSE, POWERCUTOFFREQUEST := FALSE,
       BTNEMERGENCYCUTOFF := FALSE, EMERGENCYCHAINCLOSED := TRUE, POWERCONTACTORENGAGED := FALSE);
    ADVANCE_TIME(10000000);
    fb(ENABLE := TRUE, RESET := FALSE, ARMREQUEST := FALSE, POWERCUTOFFREQUEST := FALSE,
       BTNEMERGENCYCUTOFF := FALSE, EMERGENCYCHAINCLOSED := TRUE, POWERCONTACTORENGAGED := FALSE);
    fb(ENABLE := TRUE, RESET := FALSE, ARMREQUEST := FALSE, POWERCUTOFFREQUEST := FALSE,
       BTNEMERGENCYCUTOFF := FALSE, EMERGENCYCHAINCLOSED := TRUE, POWERCONTACTORENGAGED := FALSE);
    (* 🚀 t=0 : front ArmRequest -> TestA (step 1) *)
    ADVANCE_TIME(10000000);
    fb(ENABLE := TRUE, RESET := FALSE, ARMREQUEST := TRUE, POWERCUTOFFREQUEST := FALSE,
       BTNEMERGENCYCUTOFF := FALSE, EMERGENCYCHAINCLOSED := TRUE, POWERCONTACTORENGAGED := FALSE);
    fb(ENABLE := TRUE, RESET := FALSE, ARMREQUEST := TRUE, POWERCUTOFFREQUEST := FALSE,
       BTNEMERGENCYCUTOFF := FALSE, EMERGENCYCHAINCLOSED := TRUE, POWERCONTACTORENGAGED := FALSE);
    (* 🔍 t=200ms : TestA reussi (boucle tombe) -> RestoreA *)
    ADVANCE_TIME(200000000);
    fb(ENABLE := TRUE, RESET := FALSE, ARMREQUEST := FALSE, POWERCUTOFFREQUEST := FALSE,
       BTNEMERGENCYCUTOFF := FALSE, EMERGENCYCHAINCLOSED := FALSE, POWERCONTACTORENGAGED := FALSE);
    fb(ENABLE := TRUE, RESET := FALSE, ARMREQUEST := FALSE, POWERCUTOFFREQUEST := FALSE,
       BTNEMERGENCYCUTOFF := FALSE, EMERGENCYCHAINCLOSED := FALSE, POWERCONTACTORENGAGED := FALSE);
    (* 🔍 t=400ms : RestoreA reussi -> TestB *)
    ADVANCE_TIME(200000000);
    fb(ENABLE := TRUE, RESET := FALSE, ARMREQUEST := FALSE, POWERCUTOFFREQUEST := FALSE,
       BTNEMERGENCYCUTOFF := FALSE, EMERGENCYCHAINCLOSED := TRUE, POWERCONTACTORENGAGED := FALSE);
    fb(ENABLE := TRUE, RESET := FALSE, ARMREQUEST := FALSE, POWERCUTOFFREQUEST := FALSE,
       BTNEMERGENCYCUTOFF := FALSE, EMERGENCYCHAINCLOSED := TRUE, POWERCONTACTORENGAGED := FALSE);
    (* 🔍 t=600ms : TestB reussi -> RestoreB *)
    ADVANCE_TIME(200000000);
    fb(ENABLE := TRUE, RESET := FALSE, ARMREQUEST := FALSE, POWERCUTOFFREQUEST := FALSE,
       BTNEMERGENCYCUTOFF := FALSE, EMERGENCYCHAINCLOSED := FALSE, POWERCONTACTORENGAGED := FALSE);
    fb(ENABLE := TRUE, RESET := FALSE, ARMREQUEST := FALSE, POWERCUTOFFREQUEST := FALSE,
       BTNEMERGENCYCUTOFF := FALSE, EMERGENCYCHAINCLOSED := FALSE, POWERCONTACTORENGAGED := FALSE);
    (* 🔍 t=800ms : RestoreB reussi -> PULSE (step 5), impulsion active *)
    ADVANCE_TIME(200000000);
    fb(ENABLE := TRUE, RESET := FALSE, ARMREQUEST := FALSE, POWERCUTOFFREQUEST := FALSE,
       BTNEMERGENCYCUTOFF := FALSE, EMERGENCYCHAINCLOSED := TRUE, POWERCONTACTORENGAGED := FALSE);
    fb(ENABLE := TRUE, RESET := FALSE, ARMREQUEST := FALSE, POWERCUTOFFREQUEST := FALSE,
       BTNEMERGENCYCUTOFF := FALSE, EMERGENCYCHAINCLOSED := TRUE, POWERCONTACTORENGAGED := FALSE);
    ASSERT_EQ(fb.STATUS.STATE.STEP, 5, 'precondition : pulse en cours (step 5)');
    ASSERT_TRUE(fb.CMD.ARMPULSE_CMD, 'precondition : impulsion active');

    (* ⛔ t=810ms : Enable=FALSE EN PLEINE IMPULSION -> neutralisation fail-safe (gate §2) *)
    ADVANCE_TIME(10000000);
    fb(ENABLE := FALSE, RESET := FALSE, ARMREQUEST := FALSE, POWERCUTOFFREQUEST := FALSE,
       BTNEMERGENCYCUTOFF := FALSE, EMERGENCYCHAINCLOSED := TRUE, POWERCONTACTORENGAGED := FALSE);
    fb(ENABLE := FALSE, RESET := FALSE, ARMREQUEST := FALSE, POWERCUTOFFREQUEST := FALSE,
       BTNEMERGENCYCUTOFF := FALSE, EMERGENCYCHAINCLOSED := TRUE, POWERCONTACTORENGAGED := FALSE);
    ASSERT_EQ(fb.STATUS.STATE.STEP, 0, 'Enable=FALSE -> sequence ramenee a IDLE (gate §2)');
    ASSERT_EQ(fb.STATUS.OPERATORMESSAGE, 'AU neutralisee (Enable=FALSE)', 'message neutralisation en pleine sequence (gate §2)');
    ASSERT_FALSE(fb.CMD.ARMPULSE_CMD, 'impulsion coupee immediatement (fail-safe)');
    ASSERT_FALSE(fb.CMD.MAINTAINA_CMD, 'maintien A coupe (fail-safe)');
    ASSERT_FALSE(fb.CMD.MAINTAINB_CMD, 'maintien B coupe (fail-safe)');
    ASSERT_FALSE(fb.STATUS.READY, 'Enable=FALSE -> Ready=FALSE');
    ASSERT_FALSE(fb.STATUS.DIAG.ERROR, 'neutralisation != defaut : causes repartent propres');
    ASSERT_EQ(fb.STATUS.DIAG.LASTABORTCAUSE, 0, 'neutralisation != abandon : trace repart a CST_ABORT_NONE');

    (* 🔁 t=820ms : re-Enable -> autotest repasse (boucle OK, contacteur repos) -> pret *)
    ADVANCE_TIME(10000000);
    fb(ENABLE := TRUE, RESET := FALSE, ARMREQUEST := FALSE, POWERCUTOFFREQUEST := FALSE,
       BTNEMERGENCYCUTOFF := FALSE, EMERGENCYCHAINCLOSED := TRUE, POWERCONTACTORENGAGED := FALSE);
    fb(ENABLE := TRUE, RESET := FALSE, ARMREQUEST := FALSE, POWERCUTOFFREQUEST := FALSE,
       BTNEMERGENCYCUTOFF := FALSE, EMERGENCYCHAINCLOSED := TRUE, POWERCONTACTORENGAGED := FALSE);
    ASSERT_TRUE(fb.STATUS.READY, 're-Enable sain -> Ready=TRUE (autotest repasse)');
    ASSERT_TRUE(fb.STATUS.STATE.ARMABLE, 're-Enable -> Armable=TRUE (aucun etat colle)');

    (* 🚀 t=830ms : nouvel front ArmRequest -> la sequence repart proprement depuis IDLE *)
    ADVANCE_TIME(10000000);
    fb(ENABLE := TRUE, RESET := FALSE, ARMREQUEST := TRUE, POWERCUTOFFREQUEST := FALSE,
       BTNEMERGENCYCUTOFF := FALSE, EMERGENCYCHAINCLOSED := TRUE, POWERCONTACTORENGAGED := FALSE);
    fb(ENABLE := TRUE, RESET := FALSE, ARMREQUEST := TRUE, POWERCUTOFFREQUEST := FALSE,
       BTNEMERGENCYCUTOFF := FALSE, EMERGENCYCHAINCLOSED := TRUE, POWERCONTACTORENGAGED := FALSE);
    ASSERT_EQ(fb.STATUS.STATE.STEP, 1, 'nouveau front ArmRequest -> TestA relance (retour arriere propre)');
END_TEST

TEST 'TC-P01-022 Messages par etape : branches CASE transitoires RESTORE_A/B (refermeture anticipee)'
    (* 💤 Setup : demarrage + regime etabli, sain *)
    fb(ENABLE := TRUE, RESET := FALSE, ARMREQUEST := FALSE, POWERCUTOFFREQUEST := FALSE,
       BTNEMERGENCYCUTOFF := FALSE, EMERGENCYCHAINCLOSED := TRUE, POWERCONTACTORENGAGED := FALSE);
    fb(ENABLE := TRUE, RESET := FALSE, ARMREQUEST := FALSE, POWERCUTOFFREQUEST := FALSE,
       BTNEMERGENCYCUTOFF := FALSE, EMERGENCYCHAINCLOSED := TRUE, POWERCONTACTORENGAGED := FALSE);
    ADVANCE_TIME(10000000);
    fb(ENABLE := TRUE, RESET := FALSE, ARMREQUEST := FALSE, POWERCUTOFFREQUEST := FALSE,
       BTNEMERGENCYCUTOFF := FALSE, EMERGENCYCHAINCLOSED := TRUE, POWERCONTACTORENGAGED := FALSE);
    fb(ENABLE := TRUE, RESET := FALSE, ARMREQUEST := FALSE, POWERCUTOFFREQUEST := FALSE,
       BTNEMERGENCYCUTOFF := FALSE, EMERGENCYCHAINCLOSED := TRUE, POWERCONTACTORENGAGED := FALSE);
    ASSERT_EQ(fb.STATUS.OPERATORMESSAGE, 'AU: repos - pret a rearmer', 'message CASE 0/IDLE au repos');

    (* 🚀 t=0 : front ArmRequest -> TEST_A *)
    ADVANCE_TIME(10000000);
    fb(ENABLE := TRUE, RESET := FALSE, ARMREQUEST := TRUE, POWERCUTOFFREQUEST := FALSE,
       BTNEMERGENCYCUTOFF := FALSE, EMERGENCYCHAINCLOSED := TRUE, POWERCONTACTORENGAGED := FALSE);
    fb(ENABLE := TRUE, RESET := FALSE, ARMREQUEST := TRUE, POWERCUTOFFREQUEST := FALSE,
       BTNEMERGENCYCUTOFF := FALSE, EMERGENCYCHAINCLOSED := TRUE, POWERCONTACTORENGAGED := FALSE);
    ASSERT_EQ(fb.STATUS.STATE.STEP, 1, 'TEST_A');
    ASSERT_EQ(fb.STATUS.OPERATORMESSAGE, 'AU: autotest canal A en cours', 'message CASE 1/TEST_A');

    (* 🔍 t=200ms : boucle tombe -> RESTORE_A *)
    ADVANCE_TIME(200000000);
    fb(ENABLE := TRUE, RESET := FALSE, ARMREQUEST := FALSE, POWERCUTOFFREQUEST := FALSE,
       BTNEMERGENCYCUTOFF := FALSE, EMERGENCYCHAINCLOSED := FALSE, POWERCONTACTORENGAGED := FALSE);
    fb(ENABLE := TRUE, RESET := FALSE, ARMREQUEST := FALSE, POWERCUTOFFREQUEST := FALSE,
       BTNEMERGENCYCUTOFF := FALSE, EMERGENCYCHAINCLOSED := FALSE, POWERCONTACTORENGAGED := FALSE);
    ASSERT_EQ(fb.STATUS.STATE.STEP, 2, 'RESTORE_A');
    ASSERT_EQ(fb.STATUS.OPERATORMESSAGE, 'AU: boucle urgence ouverte - verifier coup-de-poing', 'priorite §11 : boucle ouverte pendant le test A delibere');

    (* ⭐ t=250ms : refermeture ANTICIPEE (timer restore 200ms non ecoule) -> branche transitoire CASE 2 *)
    ADVANCE_TIME(50000000);
    fb(ENABLE := TRUE, RESET := FALSE, ARMREQUEST := FALSE, POWERCUTOFFREQUEST := FALSE,
       BTNEMERGENCYCUTOFF := FALSE, EMERGENCYCHAINCLOSED := TRUE, POWERCONTACTORENGAGED := FALSE);
    fb(ENABLE := TRUE, RESET := FALSE, ARMREQUEST := FALSE, POWERCUTOFFREQUEST := FALSE,
       BTNEMERGENCYCUTOFF := FALSE, EMERGENCYCHAINCLOSED := TRUE, POWERCONTACTORENGAGED := FALSE);
    ASSERT_EQ(fb.STATUS.STATE.STEP, 2, 'refermeture anticipee : toujours RESTORE_A (timer non ecoule)');
    ASSERT_EQ(fb.STATUS.OPERATORMESSAGE, 'AU: restauration canal A', 'message CASE 2/RESTORE_A (branche transitoire)');

    (* 🔍 t=400ms : timer restore termine -> TEST_B *)
    ADVANCE_TIME(150000000);
    fb(ENABLE := TRUE, RESET := FALSE, ARMREQUEST := FALSE, POWERCUTOFFREQUEST := FALSE,
       BTNEMERGENCYCUTOFF := FALSE, EMERGENCYCHAINCLOSED := TRUE, POWERCONTACTORENGAGED := FALSE);
    fb(ENABLE := TRUE, RESET := FALSE, ARMREQUEST := FALSE, POWERCUTOFFREQUEST := FALSE,
       BTNEMERGENCYCUTOFF := FALSE, EMERGENCYCHAINCLOSED := TRUE, POWERCONTACTORENGAGED := FALSE);
    ASSERT_EQ(fb.STATUS.STATE.STEP, 3, 'TEST_B');
    ASSERT_EQ(fb.STATUS.OPERATORMESSAGE, 'AU: autotest canal B en cours', 'message CASE 3/TEST_B');

    (* 🔍 t=600ms : boucle tombe -> RESTORE_B *)
    ADVANCE_TIME(200000000);
    fb(ENABLE := TRUE, RESET := FALSE, ARMREQUEST := FALSE, POWERCUTOFFREQUEST := FALSE,
       BTNEMERGENCYCUTOFF := FALSE, EMERGENCYCHAINCLOSED := FALSE, POWERCONTACTORENGAGED := FALSE);
    fb(ENABLE := TRUE, RESET := FALSE, ARMREQUEST := FALSE, POWERCUTOFFREQUEST := FALSE,
       BTNEMERGENCYCUTOFF := FALSE, EMERGENCYCHAINCLOSED := FALSE, POWERCONTACTORENGAGED := FALSE);
    ASSERT_EQ(fb.STATUS.STATE.STEP, 4, 'RESTORE_B');

    (* ⭐ t=650ms : refermeture ANTICIPEE -> branche transitoire CASE 4 *)
    ADVANCE_TIME(50000000);
    fb(ENABLE := TRUE, RESET := FALSE, ARMREQUEST := FALSE, POWERCUTOFFREQUEST := FALSE,
       BTNEMERGENCYCUTOFF := FALSE, EMERGENCYCHAINCLOSED := TRUE, POWERCONTACTORENGAGED := FALSE);
    fb(ENABLE := TRUE, RESET := FALSE, ARMREQUEST := FALSE, POWERCUTOFFREQUEST := FALSE,
       BTNEMERGENCYCUTOFF := FALSE, EMERGENCYCHAINCLOSED := TRUE, POWERCONTACTORENGAGED := FALSE);
    ASSERT_EQ(fb.STATUS.STATE.STEP, 4, 'refermeture anticipee : toujours RESTORE_B');
    ASSERT_EQ(fb.STATUS.OPERATORMESSAGE, 'AU: restauration canal B', 'message CASE 4/RESTORE_B (branche transitoire)');

    (* ⚡ t=800ms : timer restore termine -> PULSE *)
    ADVANCE_TIME(150000000);
    fb(ENABLE := TRUE, RESET := FALSE, ARMREQUEST := FALSE, POWERCUTOFFREQUEST := FALSE,
       BTNEMERGENCYCUTOFF := FALSE, EMERGENCYCHAINCLOSED := TRUE, POWERCONTACTORENGAGED := FALSE);
    fb(ENABLE := TRUE, RESET := FALSE, ARMREQUEST := FALSE, POWERCUTOFFREQUEST := FALSE,
       BTNEMERGENCYCUTOFF := FALSE, EMERGENCYCHAINCLOSED := TRUE, POWERCONTACTORENGAGED := FALSE);
    ASSERT_EQ(fb.STATUS.STATE.STEP, 5, 'PULSE');
    ASSERT_EQ(fb.STATUS.OPERATORMESSAGE, 'AU: impulsion rearmement contacteur', 'message CASE 5/PULSE');

    (* ⏱️ t=1.8s : fin d'impulsion -> CONFIRM *)
    ADVANCE_TIME(1000000000);
    fb(ENABLE := TRUE, RESET := FALSE, ARMREQUEST := FALSE, POWERCUTOFFREQUEST := FALSE,
       BTNEMERGENCYCUTOFF := FALSE, EMERGENCYCHAINCLOSED := TRUE, POWERCONTACTORENGAGED := FALSE);
    fb(ENABLE := TRUE, RESET := FALSE, ARMREQUEST := FALSE, POWERCUTOFFREQUEST := FALSE,
       BTNEMERGENCYCUTOFF := FALSE, EMERGENCYCHAINCLOSED := TRUE, POWERCONTACTORENGAGED := FALSE);
    ASSERT_EQ(fb.STATUS.STATE.STEP, 6, 'CONFIRM');
    ASSERT_EQ(fb.STATUS.OPERATORMESSAGE, 'AU: attente confirmation contacteur', 'message CASE 6/CONFIRM');

    (* ✅ t=1.81s : contacteur confirme -> IDLE *)
    ADVANCE_TIME(10000000);
    fb(ENABLE := TRUE, RESET := FALSE, ARMREQUEST := FALSE, POWERCUTOFFREQUEST := FALSE,
       BTNEMERGENCYCUTOFF := FALSE, EMERGENCYCHAINCLOSED := TRUE, POWERCONTACTORENGAGED := TRUE);
    fb(ENABLE := TRUE, RESET := FALSE, ARMREQUEST := FALSE, POWERCUTOFFREQUEST := FALSE,
       BTNEMERGENCYCUTOFF := FALSE, EMERGENCYCHAINCLOSED := TRUE, POWERCONTACTORENGAGED := TRUE);
    ASSERT_EQ(fb.STATUS.STATE.STEP, 0, 'IDLE');
    ASSERT_EQ(fb.STATUS.OPERATORMESSAGE, 'AU: repos - pret a rearmer', 'message CASE 0/IDLE apres succes');
END_TEST
